{region 'Documentation'}
(*!
<summary>Checks A-B-C registration order, delayed observation and exactly one active child.</summary>
*)
{endregion}
FUNCTION_BLOCK Test_SerialRegistrationOrder EXTENDS OrchestrationTestBase

SUPER^();

{region 'Documentation'}
(*!
<summary>Defines this scenario independently of the subject's internal fields.</summary>
*)
{endregion}
METHOD PROTECTED ConfigureScenario
FArrayLayout := E_OrchestrationArrayLayout.Ordinary;
FChildCount := 3;
ConfigureStandardSequence();
END_METHOD

END_FUNCTION_BLOCK

(* stored: Version 1.1.0.1
   POU Test_SerialRegistrationOrder: Id {c053b2de-613c-4c82-9ef5-cbd83dd4dcbc}, SpecialFunc None
   Folder Internal: Id {ead15da1-4898-400e-8ef3-fce5e8ae92d9}
   Method ConfigureScenario: Id {7db28357-147d-4dd1-af36-1d80aaed2252} *)
